(* IEC 61131-3 sources: codesys-build/examples/frame-assembly/src/generated/types, 7 files *)

(* ---- ST_LineAlarm.st ---- *)
(*
Audible alarm command for the conveyor system startup warning.
*)
TYPE ST_LineAlarm :
STRUCT
	(* Requests the audible startup warning. *)
	Active : BOOL;
END_STRUCT
END_TYPE

(* ---- ST_LineButton.st ---- *)
(*
Pushbutton pressed state and input validity.
*)
TYPE ST_LineButton :
STRUCT
	(* FALSE until the owning PLC logic supplies a current status; FALSE on stale or unavailable inputs. *)
	Valid : BOOL;
	(* TRUE while pressed; not an automatically repeating request. *)
	Pressed : BOOL;
END_STRUCT
END_TYPE

(* ---- ST_LineCollection.st ---- *)
(*
Collection lane capacity, occupancy count, and full status.
*)
TYPE ST_LineCollection :
STRUCT
	(* Maximum occupants; zero means not configured and must inhibit admission. *)
	Capacity : UINT;
	(* FALSE until the owning PLC logic supplies a current status; FALSE on stale or unavailable inputs. *)
	Valid : BOOL;
	(* Payloads physically confirmed in this collection lane. *)
	Count : UINT;
	(* Admission blocked by capacity or the configured full sensor. *)
	Full : BOOL;
END_STRUCT
END_TYPE

(* ---- ST_LineEstop.st ---- *)
(*
Supervisory emergency-stop indication for all conveyor and diverter movement. Motion requires a separate start after the stop is cleared.
*)
TYPE ST_LineEstop :
STRUCT
	(* FALSE until the owning PLC logic supplies a current status; FALSE on stale or unavailable inputs. *)
	Valid : BOOL;
	(* Observed global conveyor/diverter stop demand. Clearing it does not restart motion; a separate start is required. FALSE with invalid data does not indicate permission to run. *)
	Pressed : BOOL;
END_STRUCT
END_TYPE

(* ---- ST_LineLight.st ---- *)
(*
Separate green and red lamp outputs for a two-lamp stack light. PLC logic selects the indication and times red flashing for faults.
*)
TYPE ST_LineLight :
STRUCT
	(* Switches the green lamp on when TRUE. *)
	Green : BOOL;
	(* Switches the red lamp on when TRUE; toggle in PLC logic to flash. *)
	Red : BOOL;
END_STRUCT
END_TYPE

(* ---- ST_LinePhotoeye.st ---- *)
(*
Detection and alarm signals from a SICK RT-P4000S02 photoelectric proximity sensor.
https://www.sick.com/media/docs/7/07/907/operating_instructions_rt_photoelectric_proximity_sensor_de_en_fr_zh_ja_it_es_pt_im0050907.pdf#page=1
*)
TYPE ST_LinePhotoeye :
STRUCT
	(* Object-detection output from SICK RT-P4000S02 pin 2 (QPNP). *)
	Detection : BOOL;
	(* Sensor alarm output from SICK RT-P4000S02 pin 4. *)
	Alarm : BOOL;
END_STRUCT
END_TYPE

(* ---- ST_LineStation.st ---- *)
(*
Operator station admission, active work, waiting queue, incoming reservations, and completed work awaiting release.
*)
TYPE ST_LineStation :
STRUCT
	(* Allow new admissions. Disabling does not erase existing work or reservations. *)
	Enabled : BOOL;
	(* Waiting plus incoming reservation slots; active work is separate. *)
	ReserveCapacity : UINT := 1;
	(* FALSE until the owning PLC logic supplies a current status; FALSE on stale or unavailable inputs. *)
	Valid : BOOL;
	(* Active work payload identity. *)
	ActiveId : STRING(80);
	(* Derived admission permission including QueueFull, enable, reservations, and transfer state. *)
	CanAcceptBin : BOOL;
	(* Work completed but still physically occupies the station until outbound admission. *)
	CompletedAwaitingRelease : BOOL;
	(* Derived from configured queue sensors; do not assume suffix _1 or _2 identifies a full sensor. *)
	QueueFull : BOOL;
	(* Incoming payloads holding a waiting slot, not yet physically arrived. *)
	ReservationCount : UINT;
	(* Physically arrived waiting payloads, excluding active work and incoming reservations. *)
	WaitingCount : UINT;
END_STRUCT
END_TYPE
